Fanuc KAREL source: KD00038.KL

PROGRAM KD00038
%NOLOCKGROUP
VAR
  I: INTEGER
  J: INTEGER
  B: BOOLEAN
  R: REAL
  S: STRING[80]
BEGIN
  CONDITION[1]:
  WHEN DIN[1] = ON DO
    SIGNAL SEMAPHORE[1]
  ENDCONDITION
END KD00038
